(* IEC 61131-3 sources: Lasal-MCP/examples/SampleSource/4_PumpControlSchemeSolution/Stations/Terminal/HMI/Class/_AccContMain (part 2) *)

  end_if;

END_FUNCTION

FUNCTION VIRTUAL GLOBAL _AccContMain::IF_WindowEnd
	VAR_INPUT
		whoami 	: ^_WHOAMI;
		pic 	: ^void;
	END_VAR

  // Alle Server beim Schließen eines Fensters zurücksetzen
  //-----------------------------------------------------------------------------------------
  if (whoami^.ima <> IMA_TOUCHEDITOR) then

    clearServers();

  end_if;

END_FUNCTION

FUNCTION GLOBAL _AccContMain::DelUsbSN
  VAR
    tmpPos         : DINT;
    tmpOwnUser     : UINT;
    pActUser       : ^t_s_User;
    tmpUserName    : ARRAY[0..AccessControl_MaxUsernameLength] of CHAR;
    tmpActUserName : ARRAY[0..AccessControl_MaxUsernameLength] of CHAR;
  END_VAR

  tmpPos            := 0;
  pActUser          := NIL;
  tmpUserName[0]    := 0;
  tmpActUserName[0] := 0;

  // Benutzername angegeben
  //-----------------------------------------------------------------------------------------
  if (StrEditUserName.GetLength()) then

    StrEditUserName.GetDataAt(pData:=#tmpUserName[0], udSize:=StrEditUserName.GetLength()+1, udAt:=0);
    StrActUser.GetDataAt(pData:=#tmpActUserName[0], udSize:=StrActUser.GetLength()+1, udAt:=0);

    // Position des Benutzers holen
    tmpPos := SearchUser(pBuffer := UsersBuffer, pUserName:=#tmpUserName[0], pUser:=NIL);
    if (tmpPos >= 0) then

      // Benutzerdaten anhand der Position holen
      pActUser := getUserToEdit(to_udint(tmpPos));
      tmpOwnUser := (StrCmp(p0:=#tmpUserName[0], x1:=sizeof(tmpUserName[0]), p2:=#tmpActUserName[0], x3:=sizeof(tmpActUserName[0])));
      if ( (pActUser <> NIL) & ((tmpOwnUser) | ((tmpOwnUser = 0) & (LoggedInWithUsb = 0))) &
         (StrLen(txt:=#pActUser^.USBSerial[0], size:=sizeof(pActUser^.USBSerial[0])) <> 0) ) then

        // Berechtigt um diesen Benutzer zu bearbeiten bzw. den eigenen Benutzer bearbeiten
        if ((pActUser^.usUserLevel < ActLevel) | (tmpOwnUser = 0)) then
          pActUser^.USBSerial[0] := 0;
          refreshUserFile();
        else
          SetMSGNr(dMSGNumber:=ERR_AUTHORITY_EDITUSER);
          InsertCmd(x0:=CMD_NEWWINDOW, x1:=AccessControl_MessageWindowNr, x2:=0);
        end_if;

      else

        SetMSGNr(dMSGNumber:=ERR_DEL_USB_SERNUM);
        InsertCmd(x0:=CMD_NEWWINDOW, x1:=AccessControl_MessageWindowNr, x2:=0);

      end_if;

    else

      SetMSGNr(dMSGNumber:=ERR_USER_NOTEXIST);
      InsertCmd(x0:=CMD_NEWWINDOW, x1:=AccessControl_MessageWindowNr, x2:=0);

    end_if;

  else

    SetMSGNr(dMSGNumber:=ERR_NO_NAME);
    InsertCmd(x0:=CMD_NEWWINDOW, x1:=AccessControl_MessageWindowNr, x2:=0);

  end_if;

END_FUNCTION

FUNCTION VIRTUAL GLOBAL _AccContMain::CopyUserFile::Write
	VAR_INPUT
		input (EAX) 	: DINT;
	END_VAR
	VAR_OUTPUT
		result (EAX) 	: DINT;
	END_VAR
  VAR
    tmpExtDriveLetter : ARRAY[0..AccessControl_MaxUserFilePathLength] of CHAR;
    tmpFileCpy        : DINT;
  END_VAR

	CopyUserFile := input;
	result := CopyUserFile;

  // Exportieren/Importieren der Benutzerdatei auf einen USB-Speicher
  //-----------------------------------------------------------------------------------------
  if (CopyUserFile <> 0) then

    // USB-Speichermedium auch angeschlossen?
    //-----------------------------------------------------------------------------------------
    if (IsCon_coDriveLetter = TRUE) then          // KaiAnd, V.2.22

      if ( (coDriveLetter.GetLength() > 0) &
           (StrEditUsbSN.GetLength() > 0) ) then  // KaiAnd, V.2.22

        tmpExtDriveLetter[0] := 0;
        coDriveLetter.GetDataAt(pData:=#tmpExtDriveLetter[0], udSize:=coDriveLetter.GetLength()+1, udAt:=0);
        StrNCpy(p0:=#tmpExtDriveLetter[AccessControl_DriveLetterLength],
                x1:=sizeof(tmpExtDriveLetter[0]),
                p2:=AccessControl_UserFile,
                x3:=sizeof(_ASCII),
                ml:=AccessControl_MaxUserFilePathLength);

        // Bestehende Datei der Benutzerdaten auf entsprechendes Laufwerk kopieren
        //-----------------------------------------------------------------------------------------
        if (CopyUserFile > 0) then
          // Exportieren der Benutzerdatei auf einen USB-Speicher
          tmpFileCpy := coFileSys.FileCopy(pSource:=AccessControl_InitDriveLetter, pDest:=#tmpExtDriveLetter[0], udOption:=0);
        elsif (CopyUserFile < 0) then
          // Importieren der Benutzerdatei von einem USB-Speicher
          tmpFileCpy := coFileSys.FileCopy(pSource:=#tmpExtDriveLetter[0], pDest:=AccessControl_InitDriveLetter, udOption:=0);
        end_if;

        // Kopieren der Benutzerdaten erfolgreich?
        if (tmpFileCpy <> 0) then
          SetMSGNr(dMSGNumber:=ERR_COPYUSERS);
          InsertCmd(x0:=CMD_NEWWINDOW, x1:=AccessControl_MessageWindowNr, x2:=0);
          LogMyText("_AccContMain::CopyUserFile::Write(): Kopieren der Benutzerdaten fehlgeschlagen" );
        elsif (CopyUserFile > 0) & (tmpFileCpy = 0) then
          SetMSGNr(dMSGNumber:=MSG_EXPORT_USERS_OK);
          InsertCmd(x0:=CMD_NEWWINDOW, x1:=AccessControl_MessageWindowNr, x2:=0);
        elsif (CopyUserFile < 0) & (tmpFileCpy = 0) then
          SetMSGNr(dMSGNumber:=MSG_IMPORT_USERS_OK);
          InsertCmd(x0:=CMD_NEWWINDOW, x1:=AccessControl_MessageWindowNr, x2:=0);
        end_if;

      else  // coDriveLetter or StrEditUsbSN with emty string
        SetMSGNr(dMSGNumber:=ERR_NO_DRIVE);
        InsertCmd(x0:=CMD_NEWWINDOW, x1:=AccessControl_MessageWindowNr, x2:=0);
      end_if;

    else  // coDriveLetter client not connected
      SetMSGNr(dMSGNumber:=ERR_NO_DRIVE);
      InsertCmd(x0:=CMD_NEWWINDOW, x1:=AccessControl_MessageWindowNr, x2:=0);
    end_if;

    // Server zurücksetzen
    CopyUserFile := 0;

  end_if;

END_FUNCTION

FUNCTION _AccContMain::closeScreen

  // Benutzer befindet sich auf einem Screen, ohne korrekte Zugangsberechtigung
  if ((bCloseScreen = true) & (bdAccessConfig.IgnoreScreenAccess = 0)) then

    // Kehre zum Start-Bildschirm zurück
    InsertCmd(x0:=CMD_NEWPICTURE, x1:=coGlobal.GetStartPicture(), x2:=0);
    bCloseScreen := false;

  end_if;

END_FUNCTION

FUNCTION GLOBAL _AccContMain::CreateAdmin
	VAR_INPUT
		pUsername 	: ^CHAR;
		pPassword 	: ^CHAR;
		usLevel 	: USINT;
	END_VAR
	VAR_OUTPUT
		bSuccessful 	: BOOL;
	END_VAR

  //Rückgabewert initialisieren
  bSuccessful := FALSE;

  if (StandardUser = NIL) then

    StandardUser$^void := coSystem.Malloc(sizeof(t_s_VKUser));
    StandardUser^.pNext := NIL;

  end_if;

  //Benutzerdaten gültig?
  if ((pUsername <> NIL) & (pPassword <> NIL) & (usLevel <> NIL)) then

    StrNCpy(p0 := #StandardUser^.User.aUsername[0],
            x1 := sizeof(StandardUser^.User.aUsername[0]),
            p2 := pUsername,
            x3 := sizeof(_ASCII),
            ml := AccessControl_MaxUsernameLength);
    StrNCpy(p0 := #StandardUser^.User.aUserPassword[0],
            x1 := sizeof(StandardUser^.User.aUserPassword[0]),
            p2 := pPassword,
            x3 := sizeof(_ASCII),
            ml := AccessControl_MaxPasswordLength);
    StandardUser^.User.usUserLevel   := usLevel;
    StandardUser^.User.udUserTimeout := 0;

    bSuccessful := true;
  end_if;

END_FUNCTION

FUNCTION VIRTUAL GLOBAL _AccContMain::IF_ChkEnable
	VAR_INPUT
		key 	: DINT;
	END_VAR
	VAR_OUTPUT
		retcode 	: BOOL;
	END_VAR

  retcode := false;

  // Zugangsebenen deaktiviert (frei zugänglich)
  //-----------------------------------------------------------------------------------------
  if (Deactivate = true) then

    retcode := true;

  // Zugangscode prüfen
  //-----------------------------------------------------------------------------------------
  elsif (ActLevel >= key) then

    retcode := true;

  end_if;

END_FUNCTION

FUNCTION _AccContMain::LogMyText
VAR_INPUT
		pLogTxt 	: ^CHAR;
	END_VAR

  VAR
    NiGive	  : CmdStruct;
    NiGet     : Results;
  END_VAR

  if ((IsCon_ccSystemLogging = True) & (pLogTxt <> NIL)) then

    NiGive.uiCmd    := 0;               // Command
    NiGive.aPara[0] := (pLogTxt)$DINT;  // pointer to text

    ccSystemLogging.NewInst(#NiGive, #NiGet);

  end_if;

END_FUNCTION
